(* IEC 61131-3 sources: STruCpp/tests/st-validation/control_flow, 14 files *)

(* ---- case_statement.st ---- *)
PROGRAM CaseTest
  VAR
    basic_result : INT;
    else_result : INT;
    range_result : INT;
    selector : INT;
  END_VAR

  (* Basic CASE *)
  selector := 2;
  CASE selector OF
    1: basic_result := 10;
    2: basic_result := 20;
    3: basic_result := 30;
  END_CASE;

  (* CASE with ELSE *)
  selector := 99;
  CASE selector OF
    1: else_result := 10;
    2: else_result := 20;
  ELSE
    else_result := -1;
  END_CASE;

  (* CASE with range *)
  selector := 5;
  CASE selector OF
    1..3: range_result := 1;
    4..6: range_result := 2;
    7..9: range_result := 3;
  ELSE
    range_result := 0;
  END_CASE;
END_PROGRAM

(* ---- exit_statement.st ---- *)
PROGRAM ExitTest
  VAR
    for_exit : INT;
    while_exit : INT;
    repeat_exit : INT;
    i : INT;
  END_VAR

  (* EXIT from FOR *)
  for_exit := 0;
  FOR i := 1 TO 100 DO
    IF i > 7 THEN EXIT; END_IF;
    for_exit := for_exit + 1;
  END_FOR;

  (* EXIT from WHILE *)
  while_exit := 0;
  i := 0;
  WHILE TRUE DO
    IF i >= 4 THEN EXIT; END_IF;
    while_exit := while_exit + 1;
    i := i + 1;
  END_WHILE;

  (* EXIT from REPEAT *)
  repeat_exit := 0;
  REPEAT
    repeat_exit := repeat_exit + 1;
    IF repeat_exit >= 3 THEN EXIT; END_IF;
  UNTIL FALSE
  END_REPEAT;
END_PROGRAM

(* ---- for_loop.st ---- *)
PROGRAM ForLoopTest
  VAR
    sum_1_to_10 : INT;
    countdown : INT;
    nested_result : INT;
    early_exit_result : INT;
    step_result : INT;
    i : INT;
    j : INT;
  END_VAR

  (* Sum 1 to 10 *)
  sum_1_to_10 := 0;
  FOR i := 1 TO 10 DO
    sum_1_to_10 := sum_1_to_10 + i;
  END_FOR;

  (* Countdown *)
  countdown := 0;
  FOR i := 10 TO 1 BY -1 DO
    countdown := countdown + 1;
  END_FOR;

  (* Nested loops *)
  nested_result := 0;
  FOR i := 1 TO 3 DO
    FOR j := 1 TO 3 DO
      nested_result := nested_result + 1;
    END_FOR;
  END_FOR;

  (* Early exit *)
  early_exit_result := 0;
  FOR i := 1 TO 100 DO
    IF i > 5 THEN EXIT; END_IF;
    early_exit_result := early_exit_result + 1;
  END_FOR;

  (* Step by 2 *)
  step_result := 0;
  FOR i := 0 TO 10 BY 2 DO
    step_result := step_result + 1;
  END_FOR;
END_PROGRAM

(* ---- if_elsif_else.st ---- *)
PROGRAM IfTest
  VAR
    simple_result : INT;
    else_result : INT;
    elsif_result : INT;
    nested_result : INT;
    x : INT;
  END_VAR

  (* Simple IF *)
  simple_result := 0;
  x := 5;
  IF x > 0 THEN
    simple_result := 1;
  END_IF;

  (* IF/ELSE *)
  IF x > 10 THEN
    else_result := 1;
  ELSE
    else_result := 2;
  END_IF;

  (* IF/ELSIF/ELSE chain *)
  IF x > 10 THEN
    elsif_result := 1;
  ELSIF x > 3 THEN
    elsif_result := 2;
  ELSIF x > 0 THEN
    elsif_result := 3;
  ELSE
    elsif_result := 4;
  END_IF;

  (* Nested IF *)
  IF x > 0 THEN
    IF x < 10 THEN
      nested_result := 1;
    ELSE
      nested_result := 2;
    END_IF;
  ELSE
    nested_result := 3;
  END_IF;
END_PROGRAM

(* ---- nested_loops.st ---- *)
PROGRAM NestedLoopTest
  VAR
    matrix_sum : INT;
    break_outer : INT;
    i : INT;
    j : INT;
  END_VAR

  (* 3x4 iteration count *)
  matrix_sum := 0;
  FOR i := 1 TO 3 DO
    FOR j := 1 TO 4 DO
      matrix_sum := matrix_sum + 1;
    END_FOR;
  END_FOR;

  (* Inner EXIT only breaks inner loop *)
  break_outer := 0;
  FOR i := 1 TO 3 DO
    FOR j := 1 TO 10 DO
      IF j > 2 THEN EXIT; END_IF;
    END_FOR;
    break_outer := break_outer + 1;
  END_FOR;
END_PROGRAM

(* ---- repeat_loop.st ---- *)
PROGRAM RepeatLoopTest
  VAR
    count_result : INT;
    executes_once : INT;
    i : INT;
  END_VAR

  (* Count to 5 *)
  count_result := 0;
  i := 0;
  REPEAT
    count_result := count_result + 1;
    i := i + 1;
  UNTIL i >= 5
  END_REPEAT;

  (* Always executes at least once *)
  executes_once := 0;
  REPEAT
    executes_once := executes_once + 1;
  UNTIL TRUE
  END_REPEAT;
END_PROGRAM

(* ---- test_case_statement.st ---- *)
TEST 'CASE selects correct branch'
  VAR uut : CaseTest; END_VAR
  uut();
  ASSERT_EQ(uut.basic_result, 20);
END_TEST

TEST 'CASE ELSE for unmatched value'
  VAR uut : CaseTest; END_VAR
  uut();
  ASSERT_EQ(uut.else_result, -1);
END_TEST

TEST 'CASE with range selects correctly'
  VAR uut : CaseTest; END_VAR
  uut();
  ASSERT_EQ(uut.range_result, 2);
END_TEST

(* ---- test_exit_statement.st ---- *)
TEST 'EXIT from FOR loop'
  VAR uut : ExitTest; END_VAR
  uut();
  ASSERT_EQ(uut.for_exit, 7);
END_TEST

TEST 'EXIT from WHILE loop'
  VAR uut : ExitTest; END_VAR
  uut();
  ASSERT_EQ(uut.while_exit, 4);
END_TEST

TEST 'EXIT from REPEAT loop'
  VAR uut : ExitTest; END_VAR
  uut();
  ASSERT_EQ(uut.repeat_exit, 3);
END_TEST

(* ---- test_for_loop.st ---- *)
TEST 'Sum 1 to 10 equals 55'
  VAR uut : ForLoopTest; END_VAR
  uut();
  ASSERT_EQ(uut.sum_1_to_10, 55);
END_TEST

TEST 'Countdown executes 10 iterations'
  VAR uut : ForLoopTest; END_VAR
  uut();
  ASSERT_EQ(uut.countdown, 10);
END_TEST

TEST 'Nested loops execute 3x3=9 times'
  VAR uut : ForLoopTest; END_VAR
  uut();
  ASSERT_EQ(uut.nested_result, 9);
END_TEST

TEST 'EXIT breaks out of loop after 5 iterations'
  VAR uut : ForLoopTest; END_VAR
  uut();
  ASSERT_EQ(uut.early_exit_result, 5);
END_TEST

TEST 'Step by 2 counts 0,2,4,6,8,10 = 6 iterations'
  VAR uut : ForLoopTest; END_VAR
  uut();
  ASSERT_EQ(uut.step_result, 6);
END_TEST

(* ---- test_if_elsif_else.st ---- *)
TEST 'Simple IF with true condition'
  VAR uut : IfTest; END_VAR
  uut();
  ASSERT_EQ(uut.simple_result, 1);
END_TEST

TEST 'IF/ELSE takes else branch'
  VAR uut : IfTest; END_VAR
  uut();
  ASSERT_EQ(uut.else_result, 2);
END_TEST

TEST 'ELSIF selects first matching branch'
  VAR uut : IfTest; END_VAR
  uut();
  ASSERT_EQ(uut.elsif_result, 2);
END_TEST

TEST 'Nested IF evaluates correctly'
  VAR uut : IfTest; END_VAR
  uut();
  ASSERT_EQ(uut.nested_result, 1);
END_TEST

(* ---- test_nested_loops.st ---- *)
TEST 'Nested FOR loops 3x4 = 12 iterations'
  VAR uut : NestedLoopTest; END_VAR
  uut();
  ASSERT_EQ(uut.matrix_sum, 12);
END_TEST

TEST 'Inner EXIT only breaks inner loop'
  VAR uut : NestedLoopTest; END_VAR
  uut();
  ASSERT_EQ(uut.break_outer, 3);
END_TEST

(* ---- test_repeat_loop.st ---- *)
TEST 'REPEAT counts to 5'
  VAR uut : RepeatLoopTest; END_VAR
  uut();
  ASSERT_EQ(uut.count_result, 5);
END_TEST

TEST 'REPEAT always executes at least once'
  VAR uut : RepeatLoopTest; END_VAR
  uut();
  ASSERT_EQ(uut.executes_once, 1);
END_TEST

(* ---- test_while_loop.st ---- *)
TEST 'WHILE counts to 5'
  VAR uut : WhileLoopTest; END_VAR
  uut();
  ASSERT_EQ(uut.count_result, 5);
END_TEST

TEST 'WHILE sums 1 to 10'
  VAR uut : WhileLoopTest; END_VAR
  uut();
  ASSERT_EQ(uut.sum_result, 55);
END_TEST

TEST 'WHILE with EXIT breaks early'
  VAR uut : WhileLoopTest; END_VAR
  uut();
  ASSERT_EQ(uut.early_exit, 3);
END_TEST

(* ---- while_loop.st ---- *)
PROGRAM WhileLoopTest
  VAR
    count_result : INT;
    sum_result : INT;
    early_exit : INT;
    i : INT;
  END_VAR

  (* Count to 5 *)
  count_result := 0;
  i := 0;
  WHILE i < 5 DO
    count_result := count_result + 1;
    i := i + 1;
  END_WHILE;

  (* Sum while condition *)
  sum_result := 0;
  i := 1;
  WHILE i <= 10 DO
    sum_result := sum_result + i;
    i := i + 1;
  END_WHILE;

  (* Early exit *)
  early_exit := 0;
  i := 0;
  WHILE i < 100 DO
    IF i >= 3 THEN EXIT; END_IF;
    early_exit := early_exit + 1;
    i := i + 1;
  END_WHILE;
END_PROGRAM
